{region 'Documentation'}
(*!
<summary>Check that IN is inside the inclusive StartTime..EndTime interval.</summary>
<description>

StartTime &gt; EndTime reports Error during active evaluation; equal bounds are
valid.

A value at or beyond 24 hours reports Error before comparison or baseline capture.

</description>
*)
{endregion}
FUNCTION_BLOCK AssertInTimespan_LTOD EXTENDS AssertionBase
VAR_INPUT
    IN : LTOD; //! Actual value checked or observed by this Assertion.
    StartTime : LTOD; //! Inclusive start of the time span; must not exceed EndTime.
    EndTime : LTOD; //! Inclusive end of the time span; must not precede StartTime.
END_VAR

SUPER^();

{region 'Documentation'}
(*!
<summary>Evaluate the typed temporal relation and report higher-priority errors first.</summary>
*)
{endregion}
METHOD PROTECTED Assert
VAR
    Message : STRING(GVL_Constants.MessageLength);
    StartTimeText : STRING(GVL_Constants.AssertionValueLength);
    EndTimeText : STRING(GVL_Constants.AssertionValueLength);
    ActualText : STRING(GVL_Constants.AssertionValueLength);
END_VAR
IF NOT EvaluationActive THEN
    RETURN;
END_IF;

IF Result = E_Result.Error THEN
    RETURN;
END_IF;

IF NOT IsTimeOfDayValid_LTOD(Value := IN) THEN
    Error(Message := 'Assertion error: IN is outside the valid LTOD range (less than 24 hours).');
    RETURN;
END_IF;

IF NOT IsTimeOfDayValid_LTOD(Value := StartTime) THEN
    Error(Message := 'Assertion error: StartTime is outside the valid LTOD range (less than 24 hours).');
    RETURN;
END_IF;

IF NOT IsTimeOfDayValid_LTOD(Value := EndTime) THEN
    Error(Message := 'Assertion error: EndTime is outside the valid LTOD range (less than 24 hours).');
    RETURN;
END_IF;

IF StartTime > EndTime THEN
    StartTimeText := LTOD_TO_STRING(StartTime);
    EndTimeText := LTOD_TO_STRING(EndTime);
    Message := CONCAT('Assertion error: start time exceeds end time. StartTime = ',
        StartTimeText);
    Message := CONCAT(Message, ', EndTime = ');
    Message := CONCAT(Message, EndTimeText);
    Message := CONCAT(Message, '.');
    Error(Message := Message);
    RETURN;
END_IF;

IF Result = E_Result.Failed THEN
    RETURN;
END_IF;

IF (IN < StartTime) OR (IN > EndTime) THEN
    StartTimeText := LTOD_TO_STRING(StartTime);
    EndTimeText := LTOD_TO_STRING(EndTime);
    ActualText := LTOD_TO_STRING(IN);
    Message := CONCAT('Assertion failed: value is outside allowed timespan. StartTime = ',
        StartTimeText);
    Message := CONCAT(Message, ', EndTime = ');
    Message := CONCAT(Message, EndTimeText);
    Message := CONCAT(Message, ', Actual = ');
    Message := CONCAT(Message, ActualText);
    Message := CONCAT(Message, '.');
    Fail(Message := Message);
    RETURN;
END_IF;

Pass();
END_METHOD

END_FUNCTION_BLOCK

(* stored: Version 1.1.0.1
   POU AssertInTimespan_LTOD: Id {6768acda-26aa-41e5-a9a3-e6ad543eb763}, SpecialFunc None
   Folder Internal: Id {9a78929d-f712-46a4-b354-79a471cd2cdb}
   Method Assert: Id {4eb32e27-a369-4095-a04c-4fe736c8ac8f} *)
